(* Logix 5000 project; controller R400_500_XLS vendor 1 type 14 code 216 rev 31.11; software revision 31.01; part 18 of 32 *)
(* tags used below, declared in another part *)
   Alarm : SINT;   // Wait 3 seconds
   bResetServiceMode : BOOL;
   Condenser : INT;
   Cycles : UDT_CYCLE[11];
   DRYING : DINT;   // Drying id number
   FC45_NextMaintDate : DINT[3];   // Next maintenance due date
   I_Pw_Tnk_Lvl_Sw_Deb : BOOL;   // Debounced pure water tank level switch (100ms)
   M : DINT[5];   // Memory Bits
   ONS_FC39 : DINT;
   ONS_FC85 : SINT;
   Run : DINT;
   Service : DINT[2];   // Unused Service Mode Memory Bit
   ServicePassword : DINT;   // Service Password
   Tmr : TIMER[107];
   washerMode : SINT;   // Washer Mode Flag 0 -> Ready; 1 -> Supervisor; 2 -> Service; 3 -> Run.
   CR2Mode : SINT;   // 0= Cycle complete dry contact 1= External pure water valve
   Current_Screen : DINT;
   CycleCounter : DINT;
   FC45_NbCycBeforeMaint : DINT;
   I_Mtr_Ovrld : BOOL;   // Motor overload
   I_Pw_Tnk_Lvl_Sw : BOOL;   // Pure water tank level switch
   I_Pw_Tnk_Sft_Lvl_Sw : BOOL;   // Pure water tank safety level switch
   I_Smp_Lvl_Hgh : BOOL;   // Sump high level switch
   I_Smp_Lvl_Lw : BOOL;   // Sump low level switch
   I_Smp_Sft_Lvl_Sw : BOOL;   // Sump safety level switch
   Load : Doors;
   NumInput : UDT_NUMERIC_INPUT[65];   // Numeric input
   Q_Chm_1 : BOOL;   // Chemical pump #1
   Q_Chm_2 : BOOL;   // Chemical pump #2
   Q_Chm_3 : BOOL;   // Chemical pump #3
   Q_Chm_4 : BOOL;   // Chemical pump #4
   Q_Cld_Wtr_Fll_Vlve : BOOL;   // Cold water sump fill valve
   Q_Drn_Cldwn_Vlve : BOOL;   // Drain cool down water valve
   Q_Dry_Fan : BOOL;   // Vapor removal fan / Drying fan
   Q_Dry_Iso_Vlve : BOOL;   // Drying Isolation Valve (Normally Closed Valve)
   Q_Ht_Wtr_Fll_Vlve : BOOL;   // Hot water sump fill valve
   Q_Pw_Fll_Vlve : BOOL;   // Pure water sump/ Tank fill valve
   Screen_Ctrl : DINT;   // PLC Screen Request
   sCycleCounter : STRING;
   SumpAlarmFillTime : DINT;
   Tpb : DINT[11];
   Unit : Hrdwre;   // Unit Configuration
(* MainProgram, continued *)

ROUTINE SRE_1_SRE_6_SERVICE_MODE   (* ladder *)
// Service mode routine
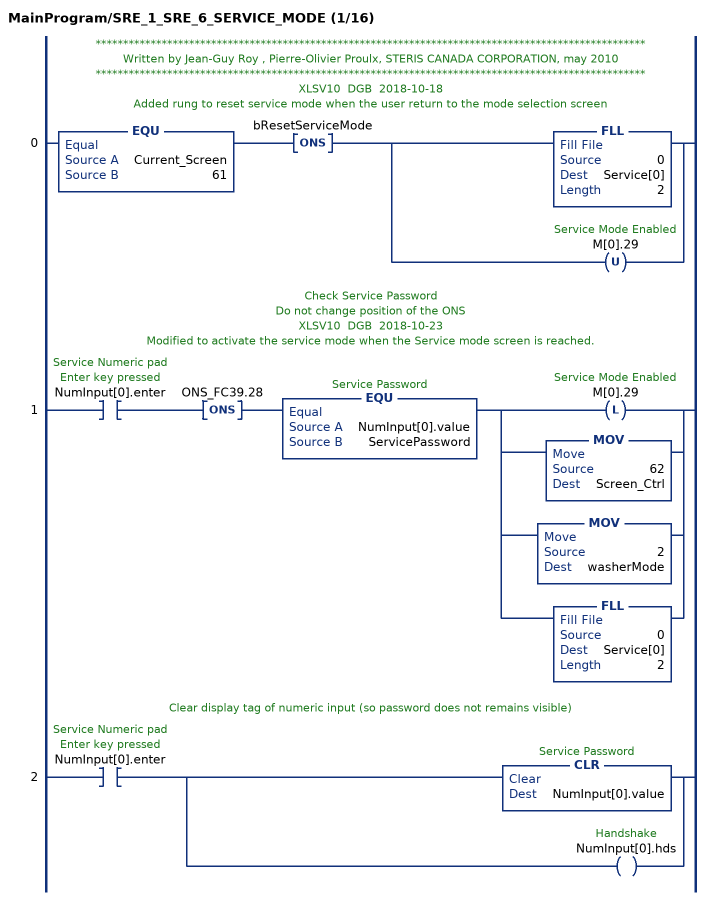
   // ****************************************************************************************************
   // Written by Jean-Guy Roy , Pierre-Olivier Proulx, STERIS CANADA CORPORATION, may 2010
   // ****************************************************************************************************
   // XLSV10  DGB  2018-10-18
   // Added rung to reset service mode when the user return to the mode selection screen
   0: EQU(Current_Screen,61)ONS(bResetServiceMode)[FLL(0,Service[0],2) ,OTU(M[0].29) ];
   // Check Service Password
   // Do not change position of the ONS
   // XLSV10  DGB  2018-10-23
   // Modified to activate the service mode when the Service mode screen is reached.
   1: XIC(NumInput[0].enter)ONS(ONS_FC39.28)EQU(NumInput[0].value,ServicePassword)[OTL(M[0].29) ,MOV(62,Screen_Ctrl) ,MOV(2,washerMode) ,FLL(0,Service[0],2) ];
   // Clear display tag of numeric input (so password does not remains visible)
   2: XIC(NumInput[0].enter)[CLR(NumInput[0].value) ,OTE(NumInput[0].hds) ];
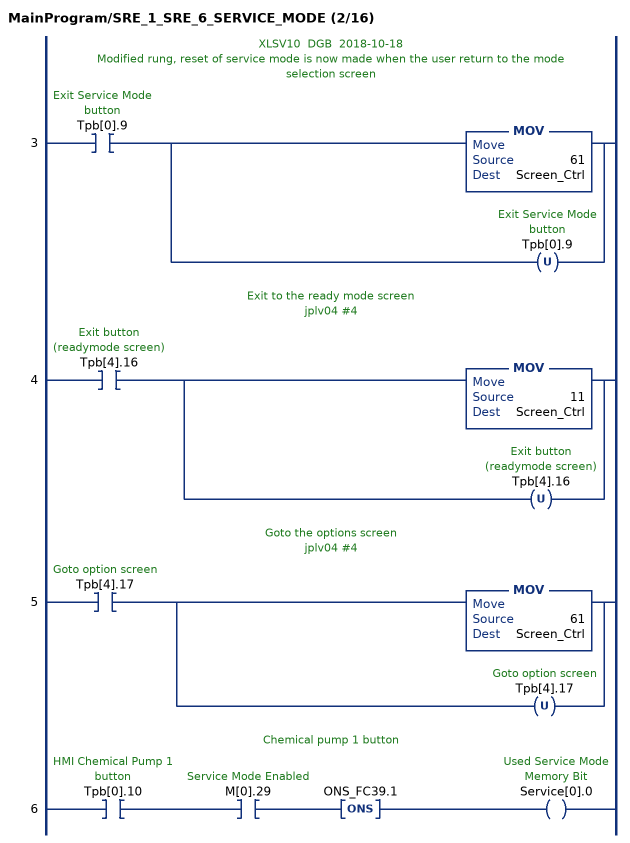
   // XLSV10  DGB  2018-10-18
   // Modified rung, reset of service mode is now made when the user return to the mode selection screen
   3: XIC(Tpb[0].9)[MOV(61,Screen_Ctrl) ,OTU(Tpb[0].9) ];
   // Exit to the ready mode screen
   // jplv04 #4
   4: XIC(Tpb[4].16)[MOV(11,Screen_Ctrl) ,OTU(Tpb[4].16) ];
   // Goto the options screen
   // jplv04 #4
   5: XIC(Tpb[4].17)[MOV(61,Screen_Ctrl) ,OTU(Tpb[4].17) ];
   // Chemical pump 1 button
   6: XIC(Tpb[0].10)XIC(M[0].29)ONS(ONS_FC39.1)OTE(Service[0].0);
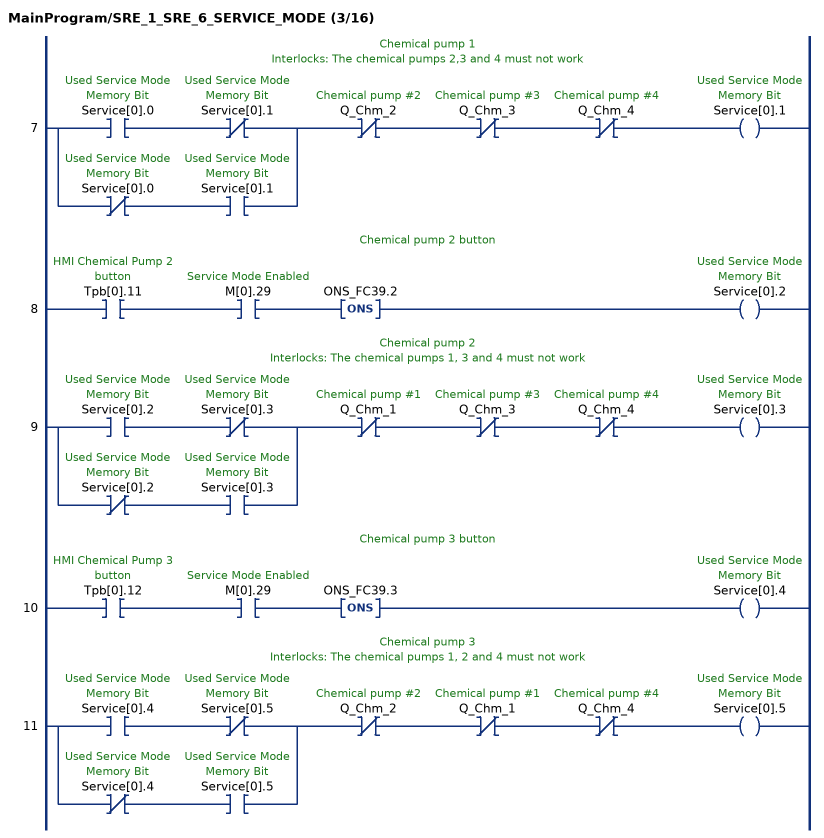
   // Chemical pump 1
   // Interlocks: The chemical pumps 2,3 and 4 must not work
   7: [XIC(Service[0].0) XIO(Service[0].1) ,XIO(Service[0].0) XIC(Service[0].1) ]XIO(Q_Chm_2)XIO(Q_Chm_3)XIO(Q_Chm_4)OTE(Service[0].1);
   // Chemical pump 2 button
   8: XIC(Tpb[0].11)XIC(M[0].29)ONS(ONS_FC39.2)OTE(Service[0].2);
   // Chemical pump 2
   // Interlocks: The chemical pumps 1, 3 and 4 must not work
   9: [XIC(Service[0].2) XIO(Service[0].3) ,XIO(Service[0].2) XIC(Service[0].3) ]XIO(Q_Chm_1)XIO(Q_Chm_3)XIO(Q_Chm_4)OTE(Service[0].3);
   // Chemical pump 3 button
   10: XIC(Tpb[0].12)XIC(M[0].29)ONS(ONS_FC39.3)OTE(Service[0].4);
   // Chemical pump 3
   // Interlocks: The chemical pumps 1, 2 and 4 must not work
   11: [XIC(Service[0].4) XIO(Service[0].5) ,XIO(Service[0].4) XIC(Service[0].5) ]XIO(Q_Chm_2)XIO(Q_Chm_1)XIO(Q_Chm_4)OTE(Service[0].5);
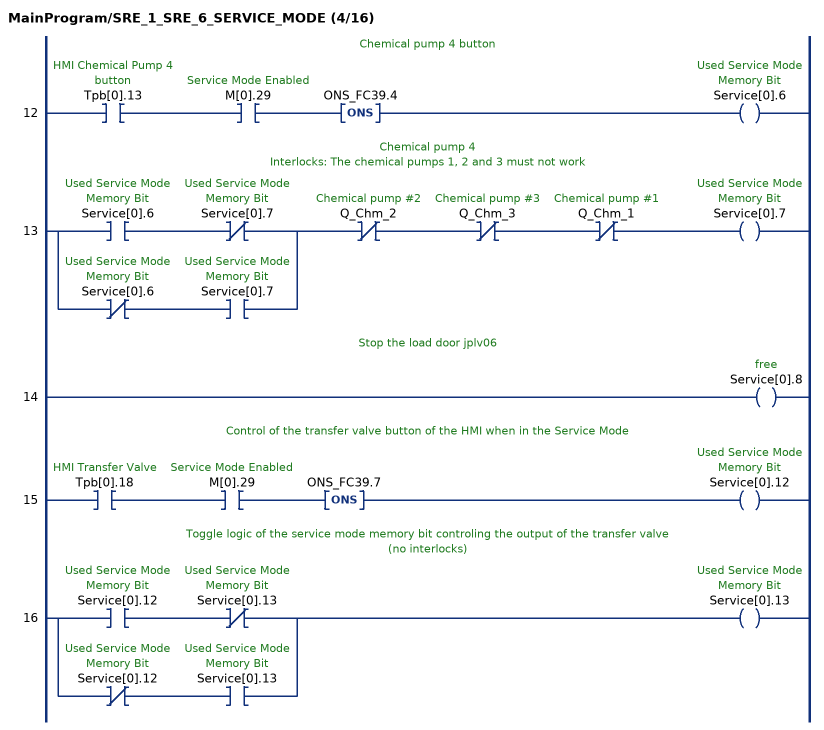
   // Chemical pump 4 button
   12: XIC(Tpb[0].13)XIC(M[0].29)ONS(ONS_FC39.4)OTE(Service[0].6);
   // Chemical pump 4
   // Interlocks: The chemical pumps 1, 2 and 3 must not work
   13: [XIC(Service[0].6) XIO(Service[0].7) ,XIO(Service[0].6) XIC(Service[0].7) ]XIO(Q_Chm_2)XIO(Q_Chm_3)XIO(Q_Chm_1)OTE(Service[0].7);
   // Stop the load door jplv06
   14: OTE(Service[0].8);
   // Control of the transfer valve button of the HMI when in the Service Mode
   15: XIC(Tpb[0].18)XIC(M[0].29)ONS(ONS_FC39.7)OTE(Service[0].12);
   // Toggle logic of the service mode memory bit controling the output of the transfer valve
   // (no interlocks)
   16: [XIC(Service[0].12) XIO(Service[0].13) ,XIO(Service[0].12) XIC(Service[0].13) ]OTE(Service[0].13);
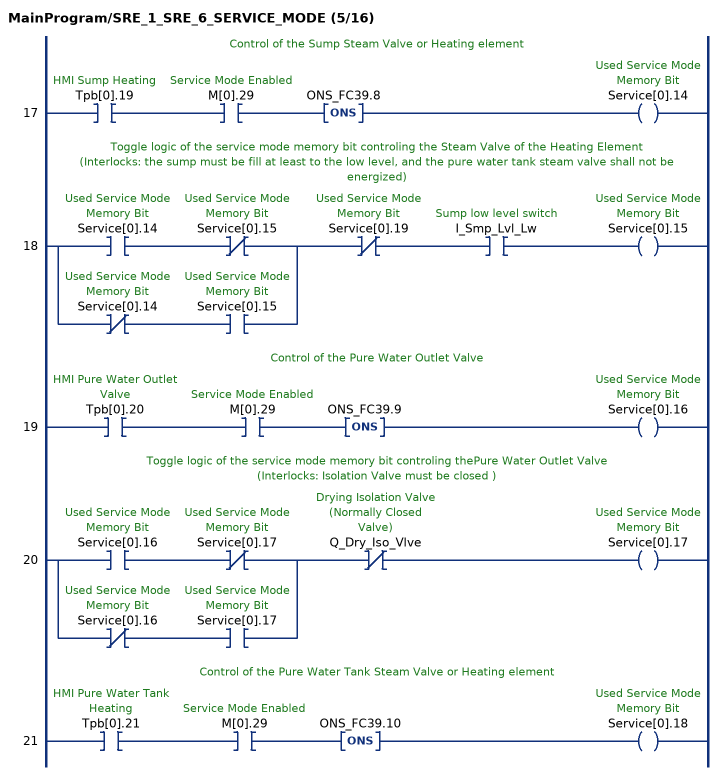
   // Control of the Sump Steam Valve or Heating element
   17: XIC(Tpb[0].19)XIC(M[0].29)ONS(ONS_FC39.8)OTE(Service[0].14);
   // Toggle logic of the service mode memory bit controling the Steam Valve of the Heating Element
   // (Interlocks: the sump must be fill at least to the low level, and the pure water tank steam valve shall not be energized)
   18: [XIC(Service[0].14) XIO(Service[0].15) ,XIO(Service[0].14) XIC(Service[0].15) ]XIO(Service[0].19)XIC(I_Smp_Lvl_Lw)OTE(Service[0].15);
   // Control of the Pure Water Outlet Valve
   19: XIC(Tpb[0].20)XIC(M[0].29)ONS(ONS_FC39.9)OTE(Service[0].16);
   // Toggle logic of the service mode memory bit controling thePure Water Outlet Valve
   // (Interlocks: Isolation Valve must be closed )
   20: [XIC(Service[0].16) XIO(Service[0].17) ,XIO(Service[0].16) XIC(Service[0].17) ]XIO(Q_Dry_Iso_Vlve)OTE(Service[0].17);
   // Control of the Pure Water Tank Steam Valve or Heating element
   21: XIC(Tpb[0].21)XIC(M[0].29)ONS(ONS_FC39.10)OTE(Service[0].18);
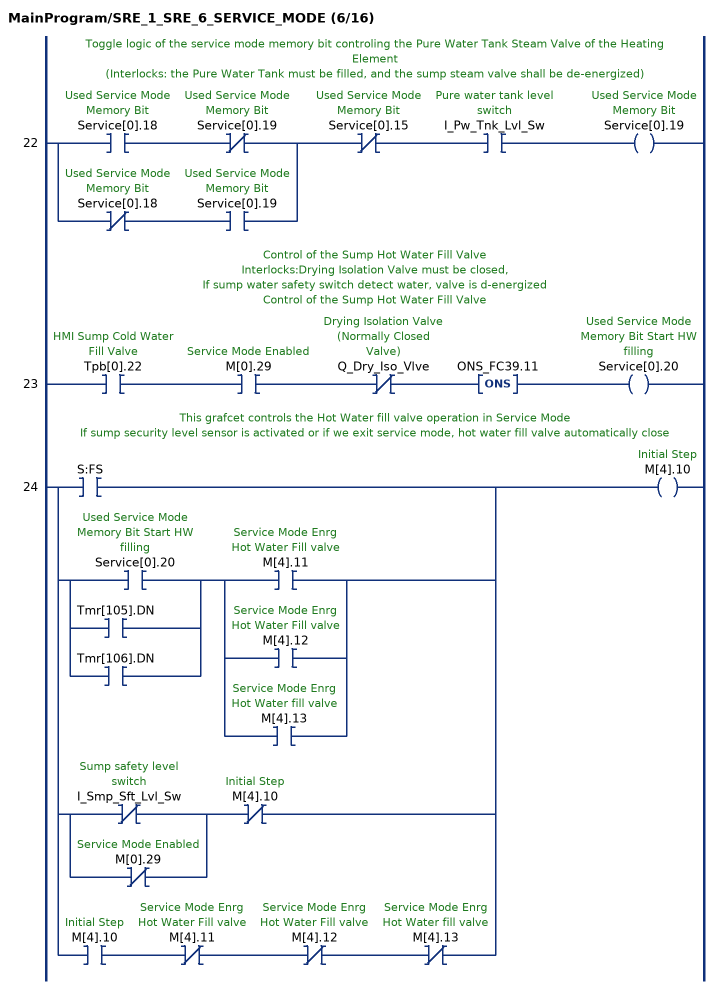
   // Toggle logic of the service mode memory bit controling the Pure Water Tank Steam Valve of the Heating Element
   // (Interlocks: the Pure Water Tank must be filled, and the sump steam valve shall be de-energized)
   22: [XIC(Service[0].18) XIO(Service[0].19) ,XIO(Service[0].18) XIC(Service[0].19) ]XIO(Service[0].15)XIC(I_Pw_Tnk_Lvl_Sw)OTE(Service[0].19);
   // Control of the Sump Hot Water Fill Valve
   // Interlocks:Drying Isolation Valve must be closed,
   // If sump water safety switch detect water, valve is d-energized
   // Control of the Sump Hot Water Fill Valve
   23: XIC(Tpb[0].22)XIC(M[0].29)XIO(Q_Dry_Iso_Vlve)ONS(ONS_FC39.11)OTE(Service[0].20);
   // This grafcet controls the Hot Water fill valve operation in Service Mode
   // If sump security level sensor is activated or if we exit service mode, hot water fill valve automatically close
   24: [XIC(S:FS) ,[XIC(Service[0].20) ,XIC(Tmr[105].DN) ,XIC(Tmr[106].DN) ] [XIC(M[4].11) ,XIC(M[4].12) ,XIC(M[4].13) ] ,[XIO(I_Smp_Sft_Lvl_Sw) ,XIO(M[0].29) ] XIO(M[4].10) ,XIC(M[4].10) XIO(M[4].11) XIO(M[4].12) XIO(M[4].13) ]OTE(M[4].10);
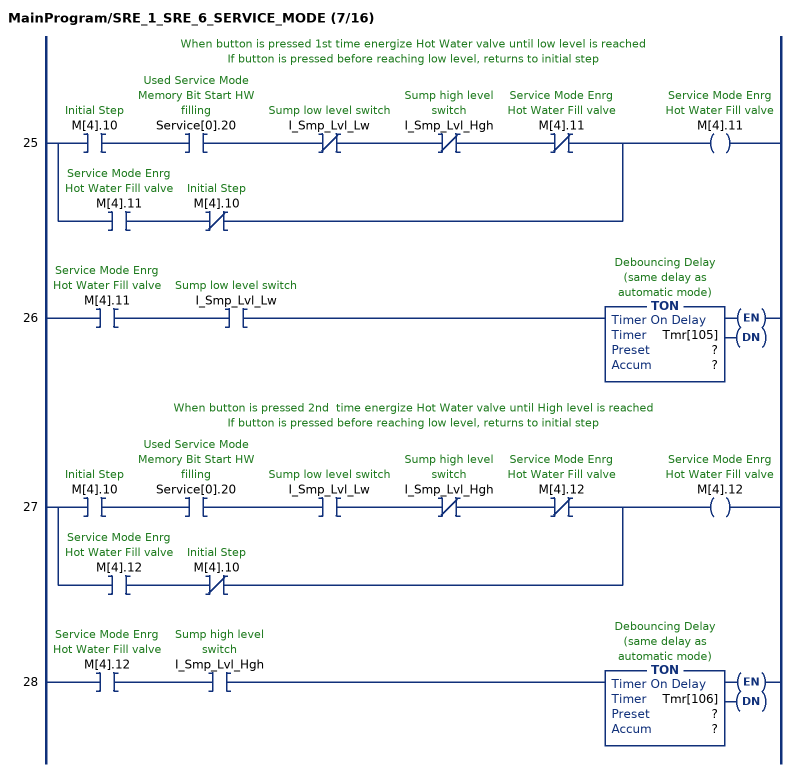
   // When button is pressed 1st time energize Hot Water valve until low level is reached
   // If button is pressed before reaching low level, returns to initial step
   25: [XIC(M[4].10) XIC(Service[0].20) XIO(I_Smp_Lvl_Lw) XIO(I_Smp_Lvl_Hgh) XIO(M[4].11) ,XIC(M[4].11) XIO(M[4].10) ]OTE(M[4].11);
   26: XIC(M[4].11)XIC(I_Smp_Lvl_Lw)TON(Tmr[105],?,?);
   // When button is pressed 2nd  time energize Hot Water valve until High level is reached
   // If button is pressed before reaching low level, returns to initial step
   27: [XIC(M[4].10) XIC(Service[0].20) XIC(I_Smp_Lvl_Lw) XIO(I_Smp_Lvl_Hgh) XIO(M[4].12) ,XIC(M[4].12) XIO(M[4].10) ]OTE(M[4].12);
   28: XIC(M[4].12)XIC(I_Smp_Lvl_Hgh)TON(Tmr[106],?,?);
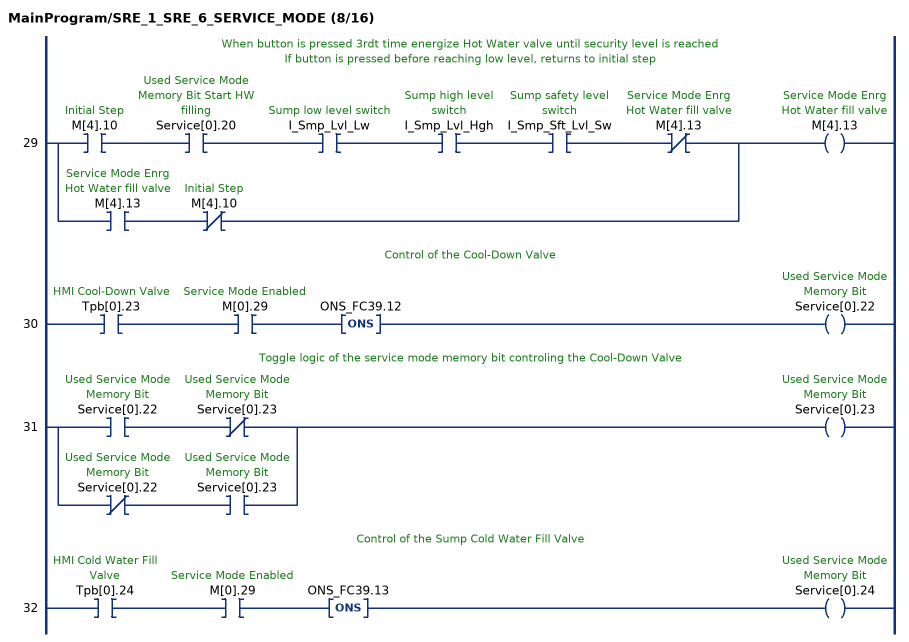
   // When button is pressed 3rdt time energize Hot Water valve until security level is reached
   // If button is pressed before reaching low level, returns to initial step
   29: [XIC(M[4].10) XIC(Service[0].20) XIC(I_Smp_Lvl_Lw) XIC(I_Smp_Lvl_Hgh) XIC(I_Smp_Sft_Lvl_Sw) XIO(M[4].13) ,XIC(M[4].13) XIO(M[4].10) ]OTE(M[4].13);
   // Control of the Cool-Down Valve
   30: XIC(Tpb[0].23)XIC(M[0].29)ONS(ONS_FC39.12)OTE(Service[0].22);
   // Toggle logic of the service mode memory bit controling the Cool-Down Valve
   31: [XIC(Service[0].22) XIO(Service[0].23) ,XIO(Service[0].22) XIC(Service[0].23) ]OTE(Service[0].23);
   // Control of the Sump Cold Water Fill Valve
   32: XIC(Tpb[0].24)XIC(M[0].29)ONS(ONS_FC39.13)OTE(Service[0].24);
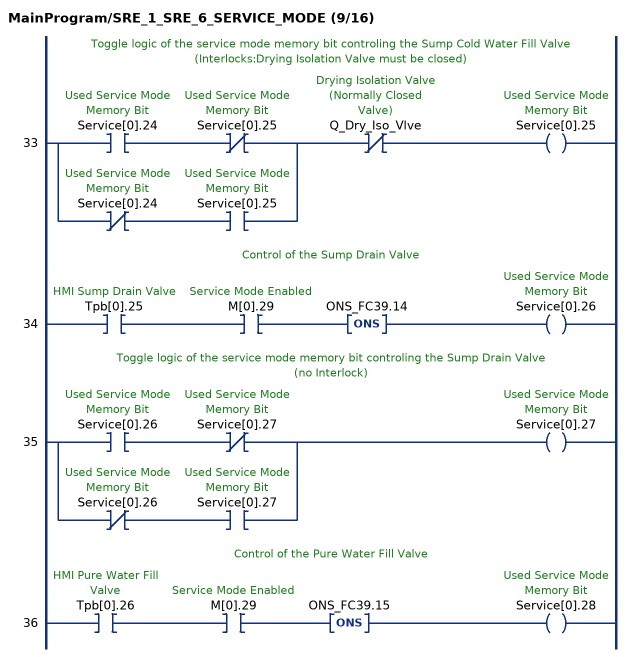
   // Toggle logic of the service mode memory bit controling the Sump Cold Water Fill Valve
   // (Interlocks:Drying Isolation Valve must be closed)
   33: [XIC(Service[0].24) XIO(Service[0].25) ,XIO(Service[0].24) XIC(Service[0].25) ]XIO(Q_Dry_Iso_Vlve)OTE(Service[0].25);
   // Control of the Sump Drain Valve
   34: XIC(Tpb[0].25)XIC(M[0].29)ONS(ONS_FC39.14)OTE(Service[0].26);
   // Toggle logic of the service mode memory bit controling the Sump Drain Valve
   // (no Interlock)
   35: [XIC(Service[0].26) XIO(Service[0].27) ,XIO(Service[0].26) XIC(Service[0].27) ]OTE(Service[0].27);
   // Control of the Pure Water Fill Valve
   36: XIC(Tpb[0].26)XIC(M[0].29)ONS(ONS_FC39.15)OTE(Service[0].28);
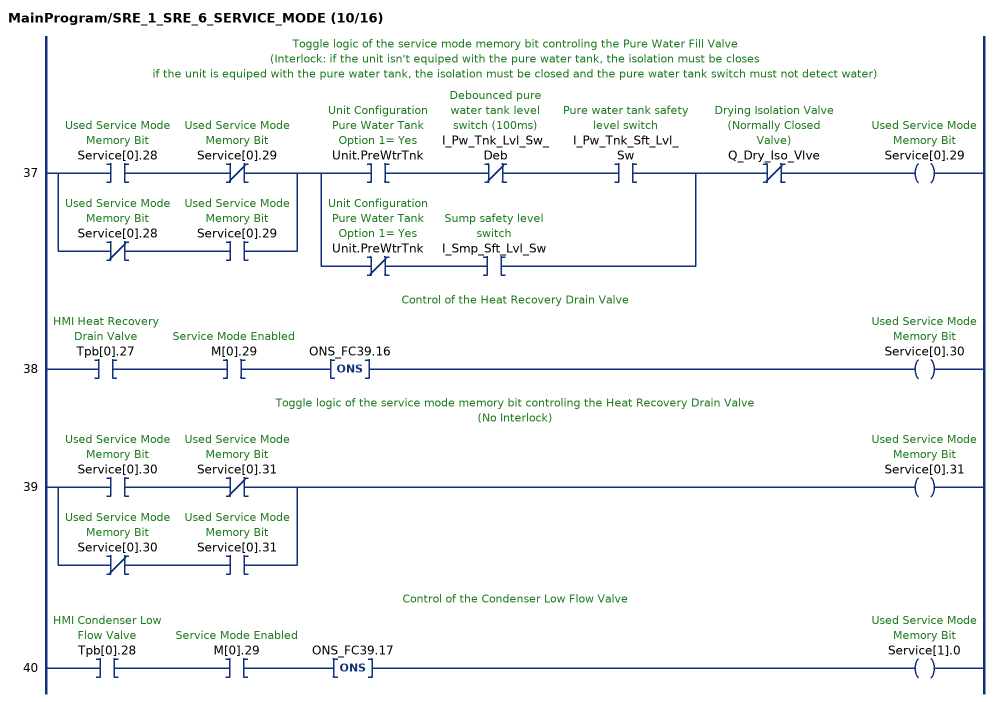
   // Toggle logic of the service mode memory bit controling the Pure Water Fill Valve
   // (Interlock: if the unit isn't equiped with the pure water tank, the isolation must be closes
   // if the unit is equiped with the pure water tank, the isolation must be closed and the pure water tank switch must not detect water)
   37: [XIC(Service[0].28) XIO(Service[0].29) ,XIO(Service[0].28) XIC(Service[0].29) ][XIC(Unit.PreWtrTnk) XIO(I_Pw_Tnk_Lvl_Sw_Deb) XIC(I_Pw_Tnk_Sft_Lvl_Sw) ,XIO(Unit.PreWtrTnk) XIC(I_Smp_Sft_Lvl_Sw) ]XIO(Q_Dry_Iso_Vlve)OTE(Service[0].29);
   // Control of the Heat Recovery Drain Valve
   38: XIC(Tpb[0].27)XIC(M[0].29)ONS(ONS_FC39.16)OTE(Service[0].30);
   // Toggle logic of the service mode memory bit controling the Heat Recovery Drain Valve
   // (No Interlock)
   39: [XIC(Service[0].30) XIO(Service[0].31) ,XIO(Service[0].30) XIC(Service[0].31) ]OTE(Service[0].31);
   // Control of the Condenser Low Flow Valve
   40: XIC(Tpb[0].28)XIC(M[0].29)ONS(ONS_FC39.17)OTE(Service[1].0);
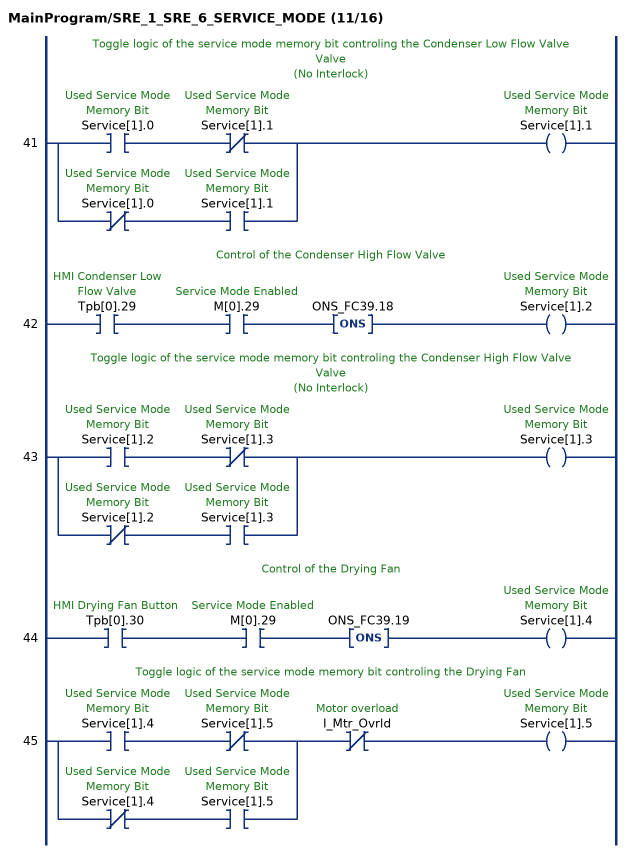
   // Toggle logic of the service mode memory bit controling the Condenser Low Flow Valve Valve
   // (No Interlock)
   41: [XIC(Service[1].0) XIO(Service[1].1) ,XIO(Service[1].0) XIC(Service[1].1) ]OTE(Service[1].1);
   // Control of the Condenser High Flow Valve
   42: XIC(Tpb[0].29)XIC(M[0].29)ONS(ONS_FC39.18)OTE(Service[1].2);
   // Toggle logic of the service mode memory bit controling the Condenser High Flow Valve Valve
   // (No Interlock)
   43: [XIC(Service[1].2) XIO(Service[1].3) ,XIO(Service[1].2) XIC(Service[1].3) ]OTE(Service[1].3);
   // Control of the Drying Fan
   44: XIC(Tpb[0].30)XIC(M[0].29)ONS(ONS_FC39.19)OTE(Service[1].4);
   // Toggle logic of the service mode memory bit controling the Drying Fan
   45: [XIC(Service[1].4) XIO(Service[1].5) ,XIO(Service[1].4) XIC(Service[1].5) ]XIO(I_Mtr_Ovrld)OTE(Service[1].5);
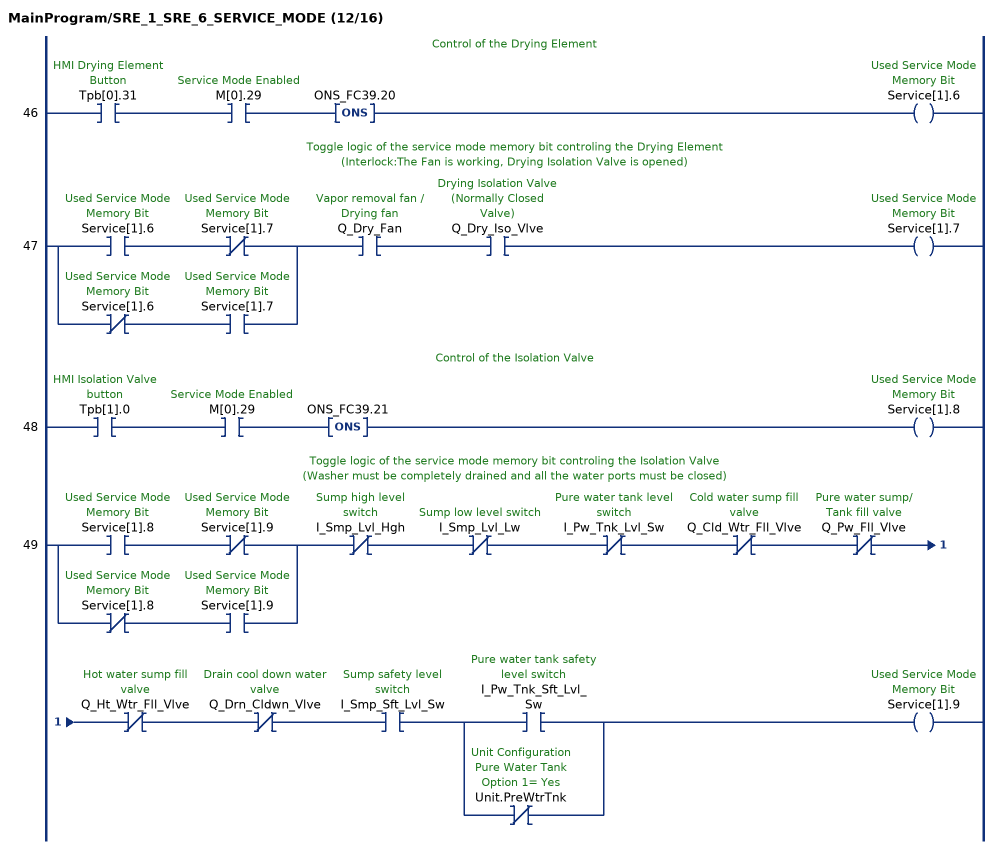
   // Control of the Drying Element
   46: XIC(Tpb[0].31)XIC(M[0].29)ONS(ONS_FC39.20)OTE(Service[1].6);
   // Toggle logic of the service mode memory bit controling the Drying Element
   // (Interlock:The Fan is working, Drying Isolation Valve is opened)
   47: [XIC(Service[1].6) XIO(Service[1].7) ,XIO(Service[1].6) XIC(Service[1].7) ]XIC(Q_Dry_Fan)XIC(Q_Dry_Iso_Vlve)OTE(Service[1].7);
   // Control of the Isolation Valve
   48: XIC(Tpb[1].0)XIC(M[0].29)ONS(ONS_FC39.21)OTE(Service[1].8);
   // Toggle logic of the service mode memory bit controling the Isolation Valve
   // (Washer must be completely drained and all the water ports must be closed)
   49: [XIC(Service[1].8) XIO(Service[1].9) ,XIO(Service[1].8) XIC(Service[1].9) ]XIO(I_Smp_Lvl_Hgh)XIO(I_Smp_Lvl_Lw)XIO(I_Pw_Tnk_Lvl_Sw)XIO(Q_Cld_Wtr_Fll_Vlve)XIO(Q_Pw_Fll_Vlve)XIO(Q_Ht_Wtr_Fll_Vlve)XIO(Q_Drn_Cldwn_Vlve)XIC(I_Smp_Sft_Lvl_Sw)[XIC(I_Pw_Tnk_Sft_Lvl_Sw) ,XIO(Unit.PreWtrTnk) ]OTE(Service[1].9);
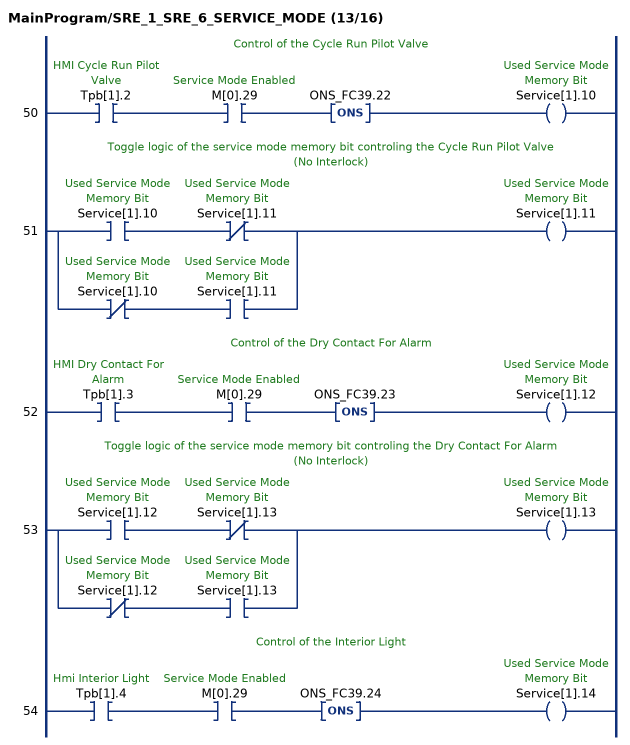
   // Control of the Cycle Run Pilot Valve
   50: XIC(Tpb[1].2)XIC(M[0].29)ONS(ONS_FC39.22)OTE(Service[1].10);
   // Toggle logic of the service mode memory bit controling the Cycle Run Pilot Valve
   // (No Interlock)
   51: [XIC(Service[1].10) XIO(Service[1].11) ,XIO(Service[1].10) XIC(Service[1].11) ]OTE(Service[1].11);
   // Control of the Dry Contact For Alarm
   52: XIC(Tpb[1].3)XIC(M[0].29)ONS(ONS_FC39.23)OTE(Service[1].12);
   // Toggle logic of the service mode memory bit controling the Dry Contact For Alarm
   // (No Interlock)
   53: [XIC(Service[1].12) XIO(Service[1].13) ,XIO(Service[1].12) XIC(Service[1].13) ]OTE(Service[1].13);
   // Control of the Interior Light
   54: XIC(Tpb[1].4)XIC(M[0].29)ONS(ONS_FC39.24)OTE(Service[1].14);
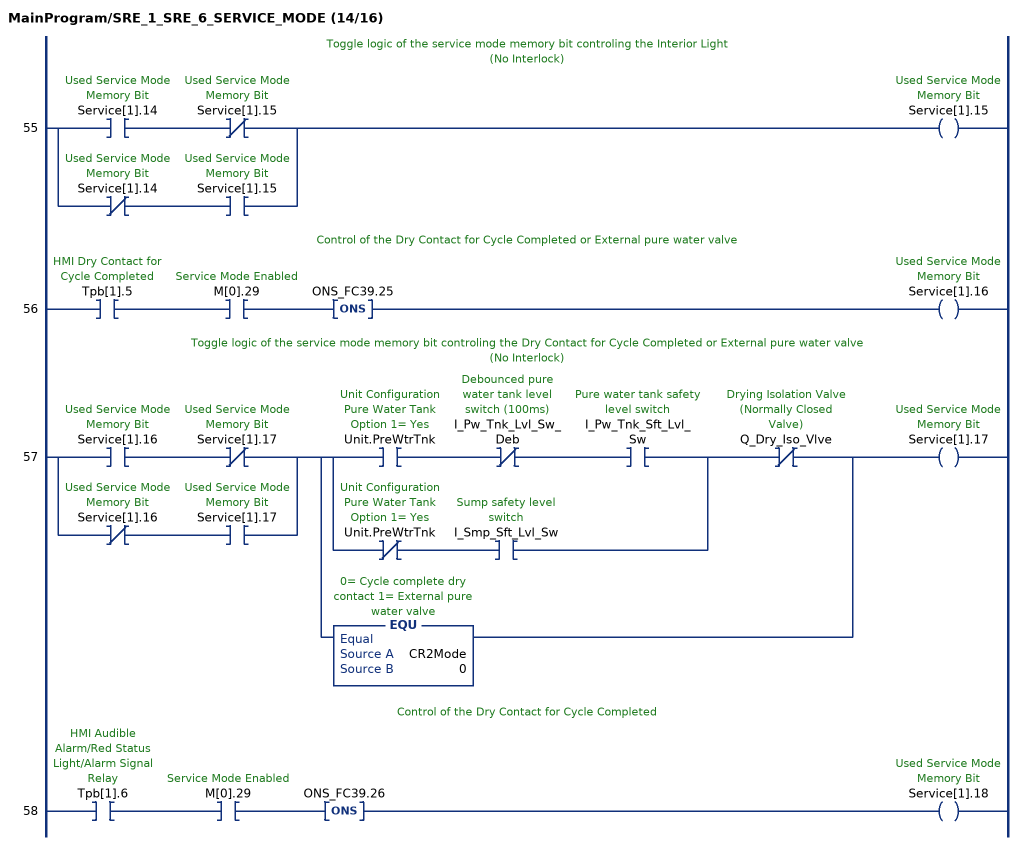
   // Toggle logic of the service mode memory bit controling the Interior Light
   // (No Interlock)
   55: [XIC(Service[1].14) XIO(Service[1].15) ,XIO(Service[1].14) XIC(Service[1].15) ]OTE(Service[1].15);
   // Control of the Dry Contact for Cycle Completed or External pure water valve
   56: XIC(Tpb[1].5)XIC(M[0].29)ONS(ONS_FC39.25)OTE(Service[1].16);
   // Toggle logic of the service mode memory bit controling the Dry Contact for Cycle Completed or External pure water valve
   // (No Interlock)
   57: [XIC(Service[1].16) XIO(Service[1].17) ,XIO(Service[1].16) XIC(Service[1].17) ][[XIC(Unit.PreWtrTnk) XIO(I_Pw_Tnk_Lvl_Sw_Deb) XIC(I_Pw_Tnk_Sft_Lvl_Sw) ,XIO(Unit.PreWtrTnk) XIC(I_Smp_Sft_Lvl_Sw) ] XIO(Q_Dry_Iso_Vlve) ,EQU(CR2Mode,0) ]OTE(Service[1].17);
   // Control of the Dry Contact for Cycle Completed
   58: XIC(Tpb[1].6)XIC(M[0].29)ONS(ONS_FC39.26)OTE(Service[1].18);
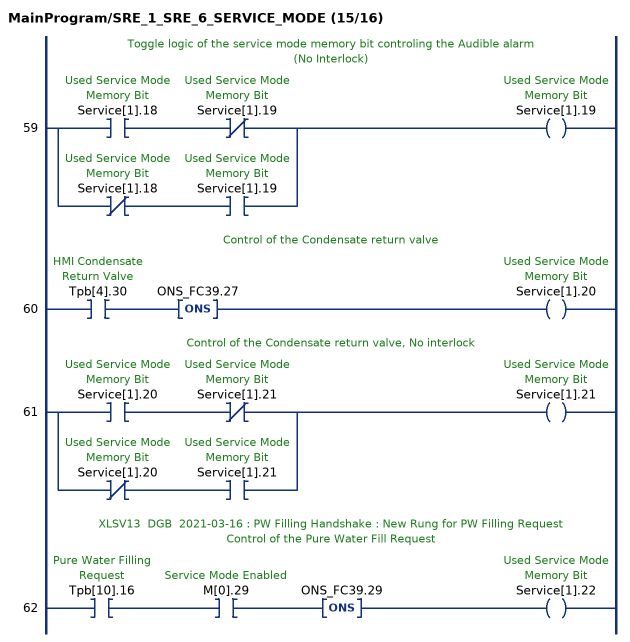
   // Toggle logic of the service mode memory bit controling the Audible alarm
   // (No Interlock)
   59: [XIC(Service[1].18) XIO(Service[1].19) ,XIO(Service[1].18) XIC(Service[1].19) ]OTE(Service[1].19);
   // Control of the Condensate return valve
   60: XIC(Tpb[4].30)ONS(ONS_FC39.27)OTE(Service[1].20);
   // Control of the Condensate return valve, No interlock
   61: [XIC(Service[1].20) XIO(Service[1].21) ,XIO(Service[1].20) XIC(Service[1].21) ]OTE(Service[1].21);
   // XLSV13  DGB  2021-03-16 : PW Filling Handshake : New Rung for PW Filling Request
   // Control of the Pure Water Fill Request
   62: XIC(Tpb[10].16)XIC(M[0].29)ONS(ONS_FC39.29)OTE(Service[1].22);
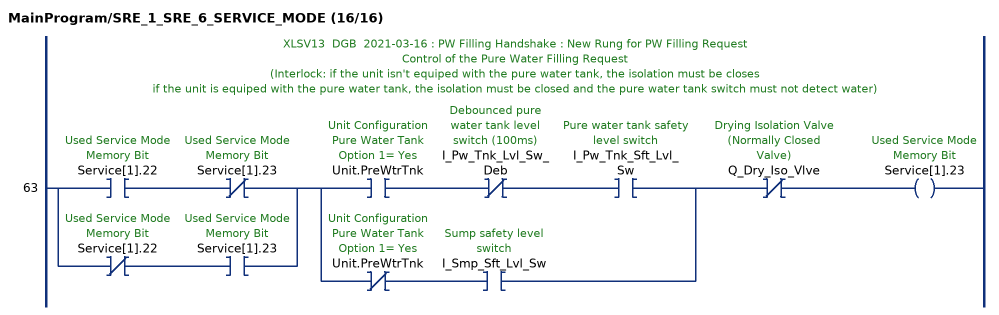
   // XLSV13  DGB  2021-03-16 : PW Filling Handshake : New Rung for PW Filling Request
   // Control of the Pure Water Filling Request
   // (Interlock: if the unit isn't equiped with the pure water tank, the isolation must be closes
   // if the unit is equiped with the pure water tank, the isolation must be closed and the pure water tank switch must not detect water)
   63: [XIC(Service[1].22) XIO(Service[1].23) ,XIO(Service[1].22) XIC(Service[1].23) ][XIC(Unit.PreWtrTnk) XIO(I_Pw_Tnk_Lvl_Sw_Deb) XIC(I_Pw_Tnk_Sft_Lvl_Sw) ,XIO(Unit.PreWtrTnk) XIC(I_Smp_Sft_Lvl_Sw) ]XIO(Q_Dry_Iso_Vlve)OTE(Service[1].23);
END_ROUTINE

ROUTINE SRE_3_HARDWARE_MACHINE_SETUP   (* ladder *)
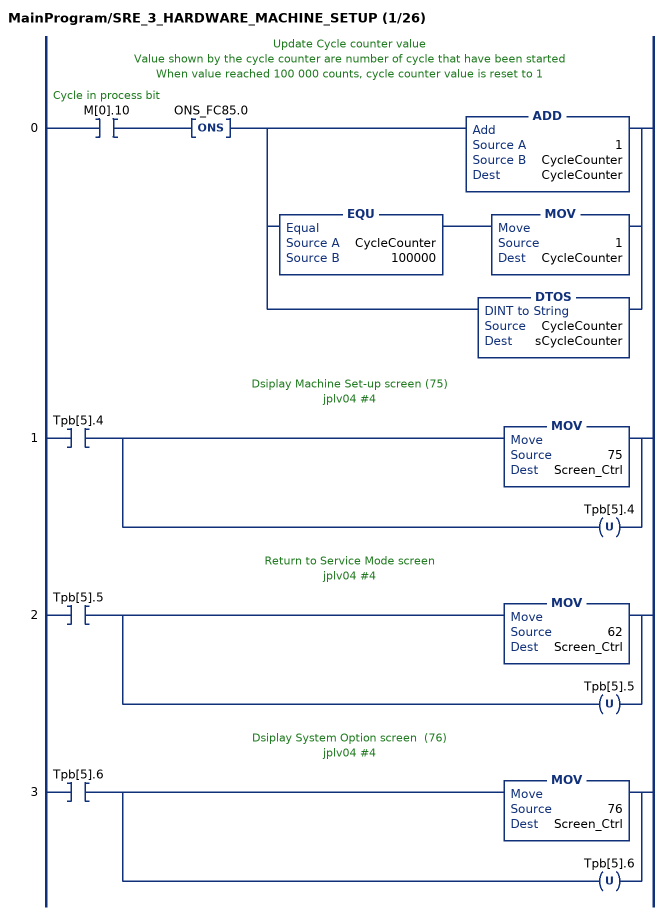
   // Update Cycle counter value
   // Value shown by the cycle counter are number of cycle that have been started
   // When value reached 100 000 counts, cycle counter value is reset to 1
   0: XIC(M[0].10)ONS(ONS_FC85.0)[ADD(1,CycleCounter,CycleCounter) ,EQU(CycleCounter,100000) MOV(1,CycleCounter) ,DTOS(CycleCounter,sCycleCounter) ];
   // Dsiplay Machine Set-up screen (75)
   // jplv04 #4
   1: XIC(Tpb[5].4)[MOV(75,Screen_Ctrl) ,OTU(Tpb[5].4) ];
   // Return to Service Mode screen
   // jplv04 #4
   2: XIC(Tpb[5].5)[MOV(62,Screen_Ctrl) ,OTU(Tpb[5].5) ];
   // Dsiplay System Option screen  (76)
   // jplv04 #4
   3: XIC(Tpb[5].6)[MOV(76,Screen_Ctrl) ,OTU(Tpb[5].6) ];
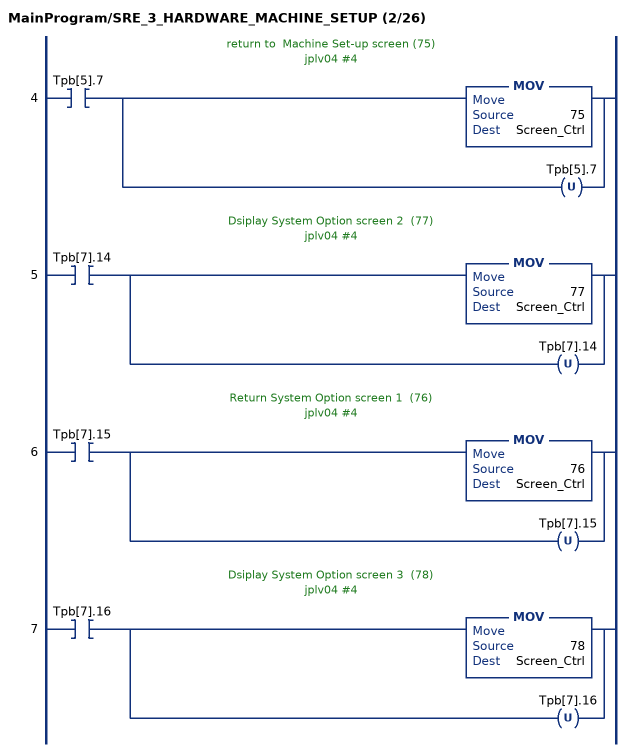
   // return to  Machine Set-up screen (75)
   // jplv04 #4
   4: XIC(Tpb[5].7)[MOV(75,Screen_Ctrl) ,OTU(Tpb[5].7) ];
   // Dsiplay System Option screen 2  (77)
   // jplv04 #4
   5: XIC(Tpb[7].14)[MOV(77,Screen_Ctrl) ,OTU(Tpb[7].14) ];
   // Return System Option screen 1  (76)
   // jplv04 #4
   6: XIC(Tpb[7].15)[MOV(76,Screen_Ctrl) ,OTU(Tpb[7].15) ];
   // Dsiplay System Option screen 3  (78)
   // jplv04 #4
   7: XIC(Tpb[7].16)[MOV(78,Screen_Ctrl) ,OTU(Tpb[7].16) ];
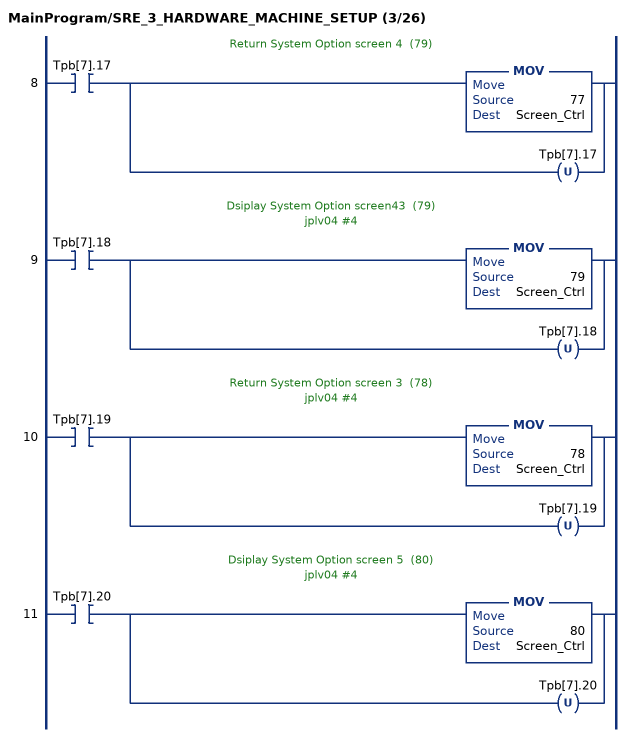
   // Return System Option screen 4  (79)
   8: XIC(Tpb[7].17)[MOV(77,Screen_Ctrl) ,OTU(Tpb[7].17) ];
   // Dsiplay System Option screen43  (79)
   // jplv04 #4
   9: XIC(Tpb[7].18)[MOV(79,Screen_Ctrl) ,OTU(Tpb[7].18) ];
   // Return System Option screen 3  (78)
   // jplv04 #4
   10: XIC(Tpb[7].19)[MOV(78,Screen_Ctrl) ,OTU(Tpb[7].19) ];
   // Dsiplay System Option screen 5  (80)
   // jplv04 #4
   11: XIC(Tpb[7].20)[MOV(80,Screen_Ctrl) ,OTU(Tpb[7].20) ];
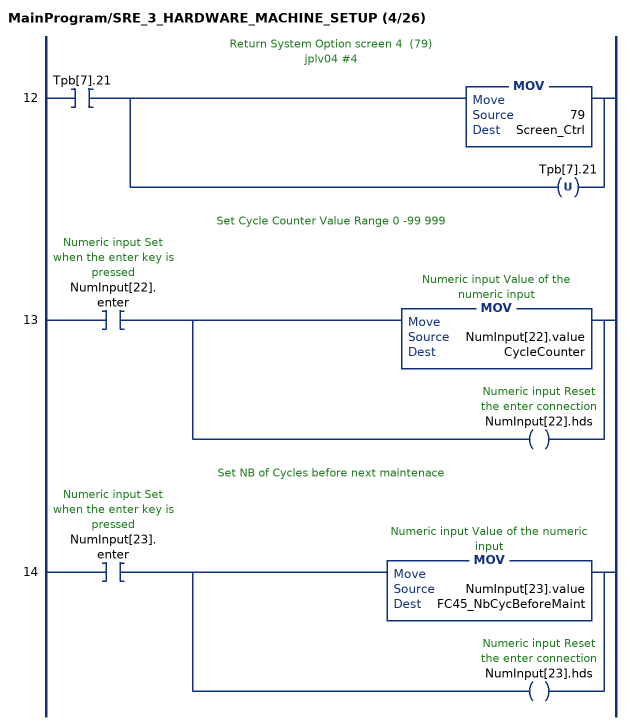
   // Return System Option screen 4  (79)
   // jplv04 #4
   12: XIC(Tpb[7].21)[MOV(79,Screen_Ctrl) ,OTU(Tpb[7].21) ];
   // Set Cycle Counter Value Range 0 -99 999
   13: XIC(NumInput[22].enter)[MOV(NumInput[22].value,CycleCounter) ,OTE(NumInput[22].hds) ];
   // Set NB of Cycles before next maintenace
   14: XIC(NumInput[23].enter)[MOV(NumInput[23].value,FC45_NbCycBeforeMaint) ,OTE(NumInput[23].hds) ];
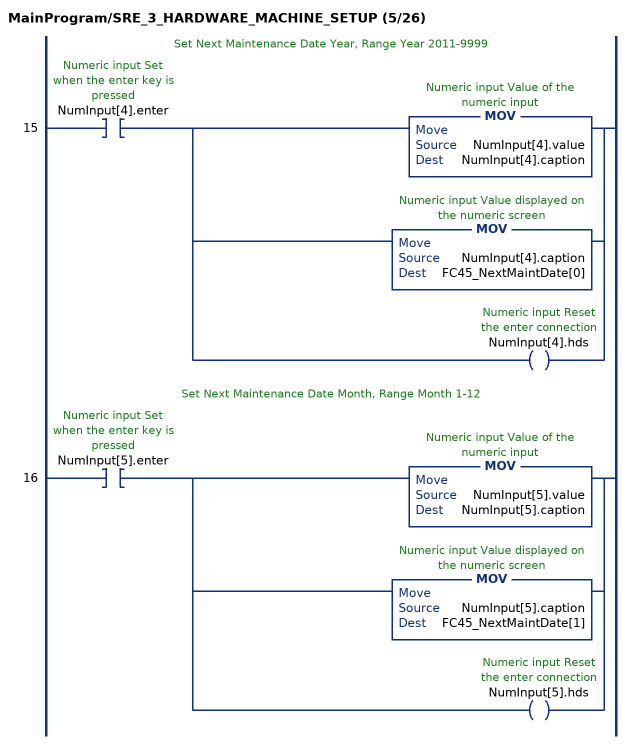
   // Set Next Maintenance Date Year, Range Year 2011-9999
   15: XIC(NumInput[4].enter)[MOV(NumInput[4].value,NumInput[4].caption) ,MOV(NumInput[4].caption,FC45_NextMaintDate[0]) ,OTE(NumInput[4].hds) ];
   // Set Next Maintenance Date Month, Range Month 1-12
   16: XIC(NumInput[5].enter)[MOV(NumInput[5].value,NumInput[5].caption) ,MOV(NumInput[5].caption,FC45_NextMaintDate[1]) ,OTE(NumInput[5].hds) ];
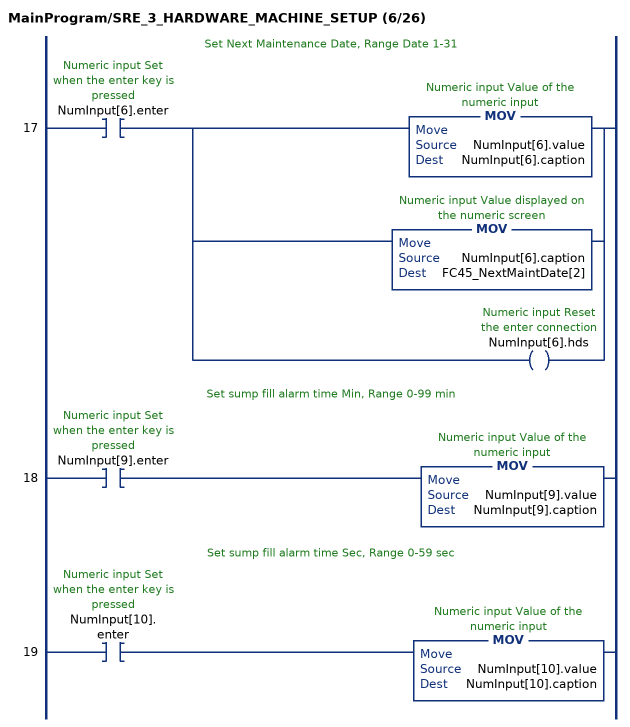
   // Set Next Maintenance Date, Range Date 1-31
   17: XIC(NumInput[6].enter)[MOV(NumInput[6].value,NumInput[6].caption) ,MOV(NumInput[6].caption,FC45_NextMaintDate[2]) ,OTE(NumInput[6].hds) ];
   // Set sump fill alarm time Min, Range 0-99 min
   18: XIC(NumInput[9].enter)MOV(NumInput[9].value,NumInput[9].caption);
   // Set sump fill alarm time Sec, Range 0-59 sec
   19: XIC(NumInput[10].enter)MOV(NumInput[10].value,NumInput[10].caption);
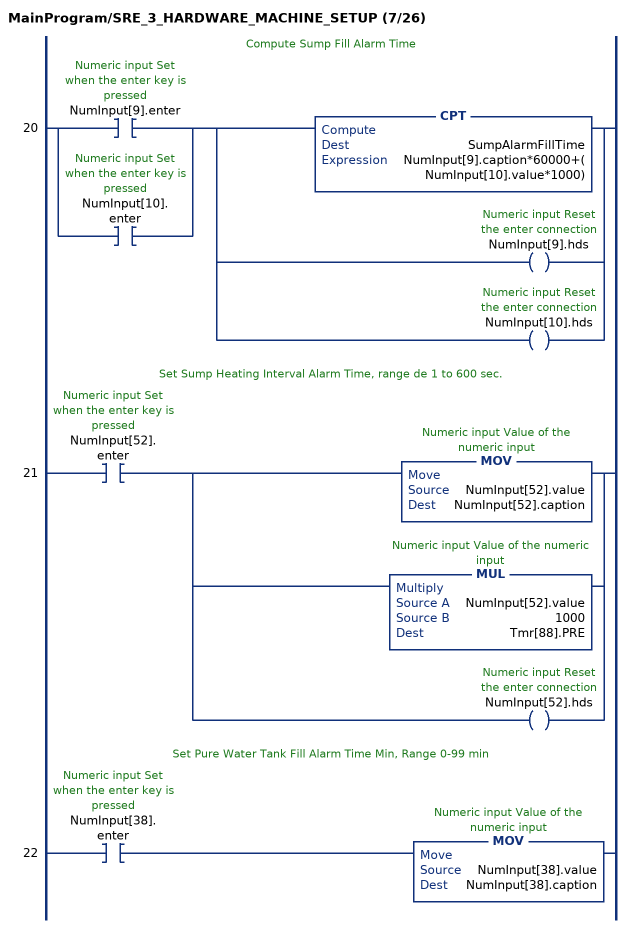
   // Compute Sump Fill Alarm Time
   20: [XIC(NumInput[9].enter) ,XIC(NumInput[10].enter) ][CPT(SumpAlarmFillTime,NumInput[9].caption*60000+(NumInput[10].value*1000)) ,OTE(NumInput[9].hds) ,OTE(NumInput[10].hds) ];
   // Set Sump Heating Interval Alarm Time, range de 1 to 600 sec.
   21: XIC(NumInput[52].enter)[MOV(NumInput[52].value,NumInput[52].caption) ,MUL(NumInput[52].value,1000,Tmr[88].PRE) ,OTE(NumInput[52].hds) ];
   // Set Pure Water Tank Fill Alarm Time Min, Range 0-99 min
   22: XIC(NumInput[38].enter)MOV(NumInput[38].value,NumInput[38].caption);
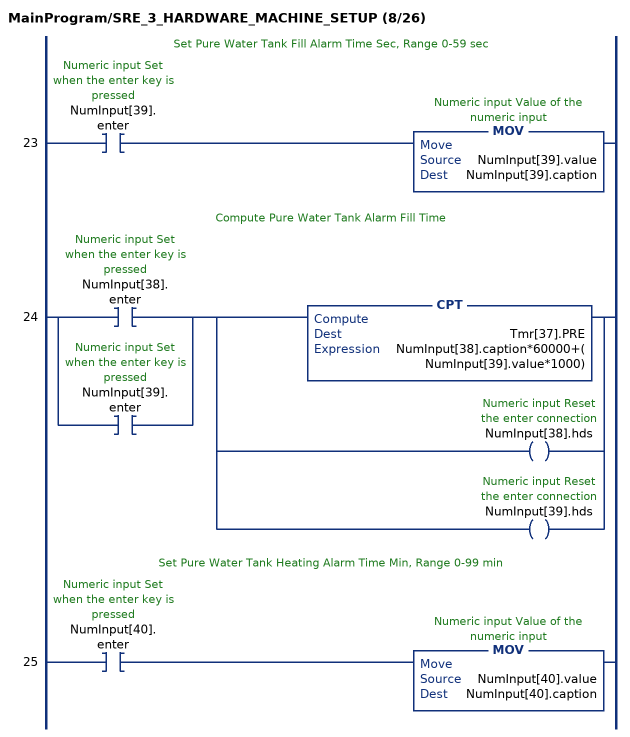
   // Set Pure Water Tank Fill Alarm Time Sec, Range 0-59 sec
   23: XIC(NumInput[39].enter)MOV(NumInput[39].value,NumInput[39].caption);
   // Compute Pure Water Tank Alarm Fill Time
   24: [XIC(NumInput[38].enter) ,XIC(NumInput[39].enter) ][CPT(Tmr[37].PRE,NumInput[38].caption*60000+(NumInput[39].value*1000)) ,OTE(NumInput[38].hds) ,OTE(NumInput[39].hds) ];
   // Set Pure Water Tank Heating Alarm Time Min, Range 0-99 min
   25: XIC(NumInput[40].enter)MOV(NumInput[40].value,NumInput[40].caption);
